Fanuc KAREL source: KD00013.KL

PROGRAM KD00013
%NOLOCKGROUP
VAR
  I: INTEGER
  J: INTEGER
  B: BOOLEAN
  R: REAL
  S: STRING[80]
BEGIN
  CLOSE HAND 1
END KD00013
